Fanuc KAREL source: KT00202.KL

PROGRAM KT00202
%NOLOCKGROUP
VAR
  I1: INTEGER
  B2: BOOLEAN
  OUT: INTEGER
BEGIN
  I1 = 2
    B2 = FALSE
  OUT = I1 AND B2
END KT00202
